SUBAPPLICATION Uebung_156_AX (* Übung zu FsWrite/FsRead: kleine Datei auf den File Server schreiben und zurücklesen *)
  (* Standard: 61499-2; Description: Copyright (c) 2026 Meisterschulen am Ostbahnhof This program and the accompanying materials are made available under the terms of the Eclipse Public License 2.0 which is available at https://www.eclipse.org/legal/epl-2.0/ SPDX-License-Identifier: EPL-2.0 *)
  (* Version 1.0, 2026-11-25, Franz Höpfinger, Meisterschulen am Ostbahnhof, initial API and implementation and/or initial documentation *)
  PACKAGE Uebungen;
  IMPORT Uebungen::const::Uebung_150_159::FileServer::FS_ADD;
  IMPORT Uebungen::const::Uebung_150_159::FileServer::FS_DATEI;
  IMPORT Uebungen::const::Uebung_150_159::FileServer::FS_FLT;
  IMPORT Uebungen::const::Uebung_150_159::FileServer::FS_TEXT;
  IMPORT isobus::pgn::ISOUSERHOME_e::network;
  IMPORT isobus::pgn::ISO_CAN_NODE::NODE1;
  IMPORT logiBUS::io::DI::logiBUS_DI::Input_I1;
  IMPORT logiBUS::io::DI::logiBUS_DI_Events::BUTTON_SINGLE_CLICK;
  IMPORT logiBUS::io::DQ::logiBUS_DO::Output_Q1;
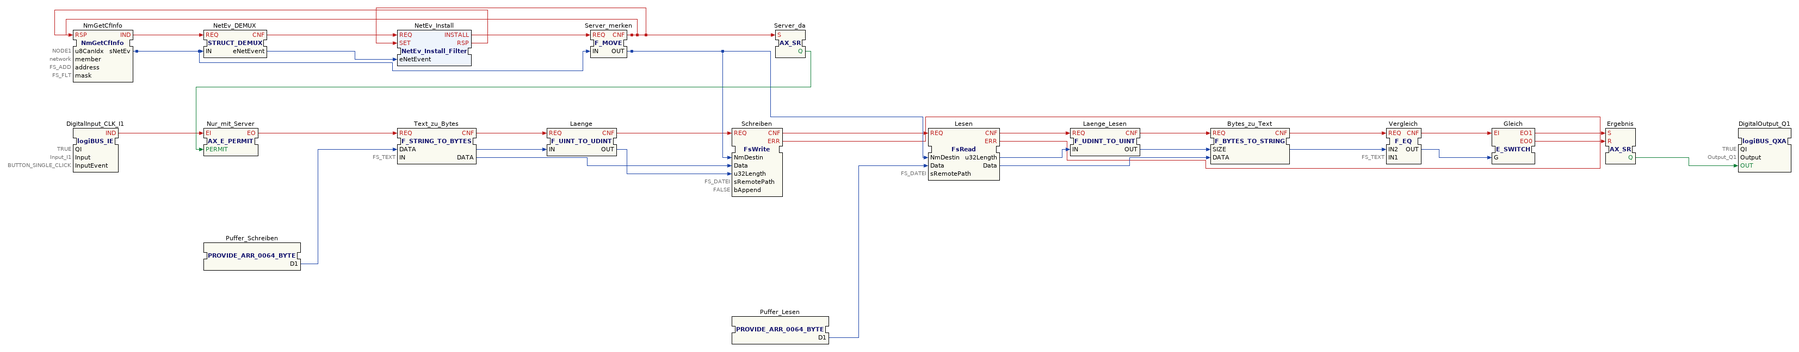
  (* File Server: Datei schreiben und zurücklesen (FsWrite, FsRead) NmGetCfInfo (network, Filter FS_ADD/FS_FLT = NAME-Funktion 61) meldet den File Server, z. B. CCI 1200 mit USB-Stick. I1 Klick (nur mit Server): FS_TEXT nach FS_DATEI schreiben, danach zurücklesen und vergleichen. Q1 an = gleich, Q1 aus = Fehler. Watch bei ERR: Schreiben/Lesen.s16Status und .u16FsError (ISO 11783-13 B.9, ab 6400 Client). FS_DATEI ohne Volume landet im aktuellen Verzeichnis des File Servers (CCI 1200: USB-Stick). Voraussetzungen: Firmware ab LOGIBUS f6afe1e4 (File Server Client), isobus_fs-ELF, PART_13_FSC = 1 in /data/functionalities.ini. Weiter: Übung 156b (FsGet/FsPut über eine lokale Datei). *)
  FBS
    NmGetCfInfo : isobus::pgn::NmGetCfInfo(u8CanIdx := NODE1, member := network, address := FS_ADD, mask := FS_FLT); (* meldet den File Server (Funktion 61) *)
    NetEv_DEMUX : eclipse4diac::convert::STRUCT_DEMUX; {SET_ATTRIBUTE(StructuredType, isobus::pgn::ISONETEVENT_T)}
    Server_merken : iec61131::selection::F_MOVE; (* eigener CF und File-Server-CF (NmDestin) *)
    Server_da : adapter::events::unidirectional::AX_SR;
    DigitalInput_CLK_I1 : logiBUS::io::DI::logiBUS_IE(QI := TRUE, Input := Input_I1, InputEvent := BUTTON_SINGLE_CLICK);
    Nur_mit_Server : adapter::events::unidirectional::AX_E_PERMIT;
    Puffer_Schreiben : eclipse4diac::convert::providers::PROVIDE_ARR_0064_BYTE;
    Text_zu_Bytes : logiBUS::utils::dyn_arr::F_STRING_TO_BYTES(IN := FS_TEXT);
    Laenge : iec61131::conversion::F_UINT_TO_UDINT;
    Schreiben : isobus::fs::FsWrite(sRemotePath := FS_DATEI, bAppend := FALSE); (* schreibt FS_TEXT nach FS_DATEI *)
    Puffer_Lesen : eclipse4diac::convert::providers::PROVIDE_ARR_0064_BYTE;
    Lesen : isobus::fs::FsRead(sRemotePath := FS_DATEI); (* liest FS_DATEI zurück *)
    Laenge_Lesen : iec61131::conversion::F_UDINT_TO_UINT;
    Bytes_zu_Text : logiBUS::utils::dyn_arr::F_BYTES_TO_STRING;
    Vergleich : iec61131::comparison::F_EQ(IN1 := FS_TEXT);
    Gleich : iec61499::events::E_SWITCH;
    Ergebnis : adapter::events::unidirectional::AX_SR; (* Q1 an = Datei gleich zurückgelesen *)
    DigitalOutput_Q1 : logiBUS::io::DQ::logiBUS_QXA(QI := TRUE, Output := Output_Q1);
  END_FBS
  SUBAPPS
    NetEv_Install : MyLib::sys::NetEv_Install_Filter;
  END_SUBAPPS
  EVENT_CONNECTIONS
    NmGetCfInfo.IND TO NetEv_DEMUX.REQ;
    NetEv_DEMUX.CNF TO NetEv_Install.REQ;
    NetEv_Install.INSTALL TO Server_merken.REQ;
    NetEv_Install.RSP TO NmGetCfInfo.RSP;
    Server_merken.CNF TO NetEv_Install.SET;
    Server_merken.CNF TO Server_da.S;
    Server_merken.CNF TO NmGetCfInfo.RSP;
    DigitalInput_CLK_I1.IND TO Nur_mit_Server.EI;
    Nur_mit_Server.EO TO Text_zu_Bytes.REQ;
    Text_zu_Bytes.CNF TO Laenge.REQ;
    Laenge.CNF TO Schreiben.REQ;
    Schreiben.CNF TO Lesen.REQ;
    Lesen.CNF TO Laenge_Lesen.REQ;
    Laenge_Lesen.CNF TO Bytes_zu_Text.REQ;
    Bytes_zu_Text.CNF TO Vergleich.REQ;
    Vergleich.CNF TO Gleich.EI;
    Gleich.EO1 TO Ergebnis.S;
    Gleich.EO0 TO Ergebnis.R;
    Schreiben.ERR TO Ergebnis.R;
    Lesen.ERR TO Ergebnis.R;
  END_CONNECTIONS
  DATA_CONNECTIONS
    NmGetCfInfo.sNetEv TO NetEv_DEMUX.IN;
    NetEv_DEMUX.eNetEvent TO NetEv_Install.eNetEvent;
    NmGetCfInfo.sNetEv TO Server_merken.IN;
    Server_merken.OUT TO Schreiben.NmDestin;
    Server_merken.OUT TO Lesen.NmDestin;
    Puffer_Schreiben.D1 TO Text_zu_Bytes.DATA;
    Text_zu_Bytes. TO Laenge.IN;
    Text_zu_Bytes.DATA TO Schreiben.Data;
    Laenge.OUT TO Schreiben.u32Length;
    Puffer_Lesen.D1 TO Lesen.Data;
    Lesen.u32Length TO Laenge_Lesen.IN;
    Laenge_Lesen.OUT TO Bytes_zu_Text.SIZE;
    Lesen.Data TO Bytes_zu_Text.DATA;
    Bytes_zu_Text. TO Vergleich.IN2;
    Vergleich.OUT TO Gleich.G;
  END_CONNECTIONS
  ADAPTER_CONNECTIONS
    Server_da.Q TO Nur_mit_Server.PERMIT;
    Ergebnis.Q TO DigitalOutput_Q1.OUT;
  END_CONNECTIONS
END_SUBAPPLICATION
